// TwinCAT 3 PLC project Untitled2
// ProgramVersion: 3.1.4026.28
// libraries:
//   Tc2_Standard, * (Beckhoff Automation GmbH)
//   Tc2_System, * (Beckhoff Automation GmbH)
// project tree:
//   DUTs/ E_PackMLStates.TcDUT
//   / PlcTask.TcTTO
//   POUs/00_System/ MAIN.TcPOU
//   POUs/01_Unit/ FB_Unit.TcPOU
//   POUs/02_Equipment/01_Palletinvoer/ FB_Palletinvoer.TcPOU, ITF_Palletinvoer.TcIO
//   POUs/02_Equipment/02_Buffer2-4/ FB_Buffer2_4.TcPOU, ITF_Buffer2_4.TcIO
//   POUs/02_Equipment/03_Buffer5/ FB_Buffer5.TcPOU, ITF_Buffer5.TcIO
//   POUs/02_Equipment/04_Depalletizer/ FB_Depalletizer.TcPOU, ITF_Depalletizer.TcIO
//   POUs/02_Equipment/05_Banddepalletizer/ FB_Banddepalletizer.TcPOU, ITF_Banddepalletizer.TcIO
//   POUs/02_Equipment/06_Palletizer/ FB_Palletizer.TcPOU, ITF_Palletizer.TcIO
//   POUs/02_Equipment/07_Blikjesband/ FB_Blikjesband.TcPOU, ITF_Blikjesband.TcIO
//   POUs/02_Equipment/08_Besturing/ FB_Besturing.TcPOU, ITF_Besturing.TcIO
//   POUs/02_Equipment/ FB_Equipment.TcPOU
//   POUs/03_Control/ FB_Control.TcPOU
//   POUs/04_Management/Alarmmanager/ FB_Alarmmanager.TcPOU
//   POUs/04_Management/HMI/ FB_HMI.TcPOU
//   POUs/04_Management/Safety/ FB_Safety.TcPOU

CONFIGURATION Untitled2
    RESOURCE PLC ON TwinCAT3
        TASK PlcTask(INTERVAL := T#10ms, PRIORITY := 20);
        PROGRAM MAIN WITH PlcTask : MAIN;
    END_RESOURCE
END_CONFIGURATION

// ---- DUTs/E_PackMLStates.TcDUT
{attribute 'qualified_only'}
{attribute 'strict'}
{attribute 'to_string'}
TYPE E_PackMLStates :
(
	Idle := 0,
	Starting, 
	Execute, 
	Suspending, 
	Suspended, 
	Unsuspending, 
	Holding,
	Held,
	Unholding,
	Resetting,
	Aborting,
	Aborted, 
	Clearing,
	Stopping,
	Stopped
);
END_TYPE

// ---- POUs/02_Equipment/01_Palletinvoer/ITF_Palletinvoer.TcIO
INTERFACE ITF_Palletinvoer

METHOD Aborted : BOOL
VAR_INPUT
END_VAR
END_METHOD

METHOD Aborting : BOOL
VAR_INPUT
END_VAR
END_METHOD

METHOD Clearing : BOOL
VAR_INPUT
END_VAR
END_METHOD

METHOD Execute : BOOL
VAR_INPUT
END_VAR
END_METHOD

METHOD Held : BOOL
VAR_INPUT
END_VAR
END_METHOD

METHOD Holding : BOOL
VAR_INPUT
END_VAR
END_METHOD

METHOD Idle : BOOL
VAR_INPUT
END_VAR
END_METHOD

METHOD Resetting : BOOL
VAR_INPUT
END_VAR
END_METHOD

METHOD Starting : BOOL
VAR_INPUT
END_VAR
END_METHOD

METHOD Stopped : BOOL
VAR_INPUT
END_VAR
END_METHOD

METHOD Stopping : BOOL
VAR_INPUT
END_VAR
END_METHOD

METHOD Suspended : BOOL
VAR_INPUT
END_VAR
END_METHOD

METHOD Suspending : BOOL
VAR_INPUT
END_VAR
END_METHOD

METHOD Unholding : BOOL
VAR_INPUT
END_VAR
END_METHOD

METHOD Unsuspending : BOOL
VAR_INPUT
END_VAR
END_METHOD

END_INTERFACE

// ---- POUs/02_Equipment/02_Buffer2-4/ITF_Buffer2_4.TcIO
INTERFACE ITF_Buffer2_4

METHOD Aborted : BOOL
VAR_INPUT
END_VAR
END_METHOD

METHOD Aborting : BOOL
VAR_INPUT
END_VAR
END_METHOD

METHOD Clearing : BOOL
VAR_INPUT
END_VAR
END_METHOD

METHOD Execute : BOOL
VAR_INPUT
END_VAR
END_METHOD

METHOD Held : BOOL
VAR_INPUT
END_VAR
END_METHOD

METHOD Holding : BOOL
VAR_INPUT
END_VAR
END_METHOD

METHOD Idle : BOOL
VAR_INPUT
END_VAR
END_METHOD

METHOD Resetting : BOOL
VAR_INPUT
END_VAR
END_METHOD

METHOD Starting : BOOL
VAR_INPUT
END_VAR
END_METHOD

METHOD Stopped : BOOL
VAR_INPUT
END_VAR
END_METHOD

METHOD Stopping : BOOL
VAR_INPUT
END_VAR
END_METHOD

METHOD Suspended : BOOL
VAR_INPUT
END_VAR
END_METHOD

METHOD Suspending : BOOL
VAR_INPUT
END_VAR
END_METHOD

METHOD Unholding : BOOL
VAR_INPUT
END_VAR
END_METHOD

METHOD Unsuspending : BOOL
VAR_INPUT
END_VAR
END_METHOD

END_INTERFACE

// ---- POUs/02_Equipment/03_Buffer5/ITF_Buffer5.TcIO
INTERFACE ITF_Buffer5

METHOD Aborted : BOOL
VAR_INPUT
END_VAR
END_METHOD

METHOD Aborting : BOOL
VAR_INPUT
END_VAR
END_METHOD

METHOD Clearing : BOOL
VAR_INPUT
END_VAR
END_METHOD

METHOD Execute : BOOL
VAR_INPUT
END_VAR
END_METHOD

METHOD Held : BOOL
VAR_INPUT
END_VAR
END_METHOD

METHOD Holding : BOOL
VAR_INPUT
END_VAR
END_METHOD

METHOD Idle : BOOL
VAR_INPUT
END_VAR
END_METHOD

METHOD Resetting : BOOL
VAR_INPUT
END_VAR
END_METHOD

METHOD Starting : BOOL
VAR_INPUT
END_VAR
END_METHOD

METHOD Stopped : BOOL
VAR_INPUT
END_VAR
END_METHOD

METHOD Stopping : BOOL
VAR_INPUT
END_VAR
END_METHOD

METHOD Suspended : BOOL
VAR_INPUT
END_VAR
END_METHOD

METHOD Suspending : BOOL
VAR_INPUT
END_VAR
END_METHOD

METHOD Unholding : BOOL
VAR_INPUT
END_VAR
END_METHOD

METHOD Unsuspending : BOOL
VAR_INPUT
END_VAR
END_METHOD

END_INTERFACE

// ---- POUs/02_Equipment/04_Depalletizer/ITF_Depalletizer.TcIO
INTERFACE ITF_Depalletizer

METHOD Aborted : BOOL
VAR_INPUT
END_VAR
END_METHOD

METHOD Aborting : BOOL
VAR_INPUT
END_VAR
END_METHOD

METHOD Clearing : BOOL
VAR_INPUT
END_VAR
END_METHOD

METHOD Execute : BOOL
VAR_INPUT
END_VAR
END_METHOD

METHOD Held : BOOL
VAR_INPUT
END_VAR
END_METHOD

METHOD Holding : BOOL
VAR_INPUT
END_VAR
END_METHOD

METHOD Idle : BOOL
VAR_INPUT
END_VAR
END_METHOD

METHOD Resetting : BOOL
VAR_INPUT
END_VAR
END_METHOD

METHOD Starting : BOOL
VAR_INPUT
END_VAR
END_METHOD

METHOD Stopped : BOOL
VAR_INPUT
END_VAR
END_METHOD

METHOD Stopping : BOOL
VAR_INPUT
END_VAR
END_METHOD

METHOD Suspended : BOOL
VAR_INPUT
END_VAR
END_METHOD

METHOD Suspending : BOOL
VAR_INPUT
END_VAR
END_METHOD

METHOD Unholding : BOOL
VAR_INPUT
END_VAR
END_METHOD

METHOD Unsuspending : BOOL
VAR_INPUT
END_VAR
END_METHOD

END_INTERFACE

// ---- POUs/02_Equipment/05_Banddepalletizer/ITF_Banddepalletizer.TcIO
INTERFACE ITF_Banddepalletizer

METHOD Aborted : BOOL
VAR_INPUT
END_VAR
END_METHOD

METHOD Aborting : BOOL
VAR_INPUT
END_VAR
END_METHOD

METHOD Clearing : BOOL
VAR_INPUT
END_VAR
END_METHOD

METHOD Execute : BOOL
VAR_INPUT
END_VAR
END_METHOD

METHOD Held : BOOL
VAR_INPUT
END_VAR
END_METHOD

METHOD Holding : BOOL
VAR_INPUT
END_VAR
END_METHOD

METHOD Idle : BOOL
VAR_INPUT
END_VAR
END_METHOD

METHOD Resetting : BOOL
VAR_INPUT
END_VAR
END_METHOD

METHOD Starting : BOOL
VAR_INPUT
END_VAR
END_METHOD

METHOD Stopped : BOOL
VAR_INPUT
END_VAR
END_METHOD

METHOD Stopping : BOOL
VAR_INPUT
END_VAR
END_METHOD

METHOD Suspended : BOOL
VAR_INPUT
END_VAR
END_METHOD

METHOD Suspending : BOOL
VAR_INPUT
END_VAR
END_METHOD

METHOD Unholding : BOOL
VAR_INPUT
END_VAR
END_METHOD

METHOD Unsuspending : BOOL
VAR_INPUT
END_VAR
END_METHOD

END_INTERFACE

// ---- POUs/02_Equipment/06_Palletizer/ITF_Palletizer.TcIO
INTERFACE ITF_Palletizer

METHOD Aborted : BOOL
VAR_INPUT
END_VAR
END_METHOD

METHOD Aborting : BOOL
VAR_INPUT
END_VAR
END_METHOD

METHOD Clearing : BOOL
VAR_INPUT
END_VAR
END_METHOD

METHOD Execute : BOOL
VAR_INPUT
END_VAR
END_METHOD

METHOD Held : BOOL
VAR_INPUT
END_VAR
END_METHOD

METHOD Holding : BOOL
VAR_INPUT
END_VAR
END_METHOD

METHOD Idle : BOOL
VAR_INPUT
END_VAR
END_METHOD

METHOD Resetting : BOOL
VAR_INPUT
END_VAR
END_METHOD

METHOD Starting : BOOL
VAR_INPUT
END_VAR
END_METHOD

METHOD Stopped : BOOL
VAR_INPUT
END_VAR
END_METHOD

METHOD Stopping : BOOL
VAR_INPUT
END_VAR
END_METHOD

METHOD Suspended : BOOL
VAR_INPUT
END_VAR
END_METHOD

METHOD Suspending : BOOL
VAR_INPUT
END_VAR
END_METHOD

METHOD Unholding : BOOL
VAR_INPUT
END_VAR
END_METHOD

METHOD Unsuspending : BOOL
VAR_INPUT
END_VAR
END_METHOD

END_INTERFACE

// ---- POUs/02_Equipment/07_Blikjesband/ITF_Blikjesband.TcIO
INTERFACE ITF_Blikjesband

METHOD Aborted : BOOL
VAR_INPUT
END_VAR
END_METHOD

METHOD Aborting : BOOL
VAR_INPUT
END_VAR
END_METHOD

METHOD Clearing : BOOL
VAR_INPUT
END_VAR
END_METHOD

METHOD Execute : BOOL
VAR_INPUT
END_VAR
END_METHOD

METHOD Held : BOOL
VAR_INPUT
END_VAR
END_METHOD

METHOD Holding : BOOL
VAR_INPUT
END_VAR
END_METHOD

METHOD Idle : BOOL
VAR_INPUT
END_VAR
END_METHOD

METHOD Resetting : BOOL
VAR_INPUT
END_VAR
END_METHOD

METHOD Starting : BOOL
VAR_INPUT
END_VAR
END_METHOD

METHOD Stopped : BOOL
VAR_INPUT
END_VAR
END_METHOD

METHOD Stopping : BOOL
VAR_INPUT
END_VAR
END_METHOD

METHOD Suspended : BOOL
VAR_INPUT
END_VAR
END_METHOD

METHOD Suspending : BOOL
VAR_INPUT
END_VAR
END_METHOD

METHOD Unholding : BOOL
VAR_INPUT
END_VAR
END_METHOD

METHOD Unsuspending : BOOL
VAR_INPUT
END_VAR
END_METHOD

END_INTERFACE

// ---- POUs/02_Equipment/08_Besturing/ITF_Besturing.TcIO
INTERFACE ITF_Besturing

METHOD StatusLampGeel : BOOL
VAR_INPUT
END_VAR
END_METHOD

METHOD StatusLampGroen : BOOL
VAR_INPUT
END_VAR
END_METHOD

METHOD StatusLampRood : BOOL
VAR_INPUT
END_VAR
END_METHOD

END_INTERFACE

// ---- POUs/00_System/MAIN.TcPOU
PROGRAM MAIN
VAR
	test : BOOL;
END_VAR

// Klopt dit?

END_PROGRAM

// ---- POUs/01_Unit/FB_Unit.TcPOU
FUNCTION_BLOCK FB_Unit
VAR_INPUT
END_VAR
VAR_OUTPUT
END_VAR
VAR
END_VAR

END_FUNCTION_BLOCK

// ---- POUs/02_Equipment/01_Palletinvoer/FB_Palletinvoer.TcPOU
FUNCTION_BLOCK FB_Palletinvoer IMPLEMENTS ITF_Palletinvoer
VAR_INPUT
END_VAR
VAR_OUTPUT
END_VAR
VAR
END_VAR

{warning 'Add method implementation '}
METHOD Aborted : BOOL
END_METHOD

{warning 'Add method implementation '}
METHOD Aborting : BOOL
END_METHOD

{warning 'Add method implementation '}
METHOD Clearing : BOOL
END_METHOD

{warning 'Add method implementation '}
METHOD Execute : BOOL
END_METHOD

{warning 'Add method implementation '}
METHOD Held : BOOL
END_METHOD

{warning 'Add method implementation '}
METHOD Holding : BOOL
END_METHOD

{warning 'Add method implementation '}
METHOD Idle : BOOL
END_METHOD

{warning 'Add method implementation '}
METHOD Resetting : BOOL
END_METHOD

{warning 'Add method implementation '}
METHOD Starting : BOOL
END_METHOD

{warning 'Add method implementation '}
METHOD Stopped : BOOL
END_METHOD

{warning 'Add method implementation '}
METHOD Stopping : BOOL
END_METHOD

{warning 'Add method implementation '}
METHOD Suspended : BOOL
END_METHOD

{warning 'Add method implementation '}
METHOD Suspending : BOOL
END_METHOD

{warning 'Add method implementation '}
METHOD Unholding : BOOL
END_METHOD

{warning 'Add method implementation '}
METHOD Unsuspending : BOOL
END_METHOD

END_FUNCTION_BLOCK

// ---- POUs/02_Equipment/02_Buffer2-4/FB_Buffer2_4.TcPOU
FUNCTION_BLOCK FB_Buffer2_4 IMPLEMENTS ITF_Buffer2_4
VAR_INPUT
END_VAR
VAR_OUTPUT
END_VAR
VAR
END_VAR

{warning 'Add method implementation '}
METHOD Aborted : BOOL
END_METHOD

{warning 'Add method implementation '}
METHOD Aborting : BOOL
END_METHOD

{warning 'Add method implementation '}
METHOD Clearing : BOOL
END_METHOD

{warning 'Add method implementation '}
METHOD Execute : BOOL
END_METHOD

{warning 'Add method implementation '}
METHOD Held : BOOL
END_METHOD

{warning 'Add method implementation '}
METHOD Holding : BOOL
END_METHOD

{warning 'Add method implementation '}
METHOD Idle : BOOL
END_METHOD

{warning 'Add method implementation '}
METHOD Resetting : BOOL
END_METHOD

{warning 'Add method implementation '}
METHOD Starting : BOOL
END_METHOD

{warning 'Add method implementation '}
METHOD Stopped : BOOL
END_METHOD

{warning 'Add method implementation '}
METHOD Stopping : BOOL
END_METHOD

{warning 'Add method implementation '}
METHOD Suspended : BOOL
END_METHOD

{warning 'Add method implementation '}
METHOD Suspending : BOOL
END_METHOD

{warning 'Add method implementation '}
METHOD Unholding : BOOL
END_METHOD

{warning 'Add method implementation '}
METHOD Unsuspending : BOOL
END_METHOD

END_FUNCTION_BLOCK

// ---- POUs/02_Equipment/03_Buffer5/FB_Buffer5.TcPOU
FUNCTION_BLOCK FB_Buffer5 IMPLEMENTS ITF_Buffer5
VAR_INPUT
END_VAR
VAR_OUTPUT
END_VAR
VAR
END_VAR

{warning 'Add method implementation '}
METHOD Aborted : BOOL
END_METHOD

{warning 'Add method implementation '}
METHOD Aborting : BOOL
END_METHOD

{warning 'Add method implementation '}
METHOD Clearing : BOOL
END_METHOD

{warning 'Add method implementation '}
METHOD Execute : BOOL
END_METHOD

{warning 'Add method implementation '}
METHOD Held : BOOL
END_METHOD

{warning 'Add method implementation '}
METHOD Holding : BOOL
END_METHOD

{warning 'Add method implementation '}
METHOD Idle : BOOL
END_METHOD

{warning 'Add method implementation '}
METHOD Resetting : BOOL
END_METHOD

{warning 'Add method implementation '}
METHOD Starting : BOOL
END_METHOD

{warning 'Add method implementation '}
METHOD Stopped : BOOL
END_METHOD

{warning 'Add method implementation '}
METHOD Stopping : BOOL
END_METHOD

{warning 'Add method implementation '}
METHOD Suspended : BOOL
END_METHOD

{warning 'Add method implementation '}
METHOD Suspending : BOOL
END_METHOD

{warning 'Add method implementation '}
METHOD Unholding : BOOL
END_METHOD

{warning 'Add method implementation '}
METHOD Unsuspending : BOOL
END_METHOD

END_FUNCTION_BLOCK

// ---- POUs/02_Equipment/04_Depalletizer/FB_Depalletizer.TcPOU
FUNCTION_BLOCK FB_Depalletizer IMPLEMENTS ITF_Depalletizer
VAR_INPUT
END_VAR
VAR_OUTPUT
END_VAR
VAR
END_VAR

{warning 'Add method implementation '}
METHOD Aborted : BOOL
END_METHOD

{warning 'Add method implementation '}
METHOD Aborting : BOOL
END_METHOD

{warning 'Add method implementation '}
METHOD Clearing : BOOL
END_METHOD

{warning 'Add method implementation '}
METHOD Execute : BOOL
END_METHOD

{warning 'Add method implementation '}
METHOD Held : BOOL
END_METHOD

{warning 'Add method implementation '}
METHOD Holding : BOOL
END_METHOD

{warning 'Add method implementation '}
METHOD Idle : BOOL
END_METHOD

{warning 'Add method implementation '}
METHOD Resetting : BOOL
END_METHOD

{warning 'Add method implementation '}
METHOD Starting : BOOL
END_METHOD

{warning 'Add method implementation '}
METHOD Stopped : BOOL
END_METHOD

{warning 'Add method implementation '}
METHOD Stopping : BOOL
END_METHOD

{warning 'Add method implementation '}
METHOD Suspended : BOOL
END_METHOD

{warning 'Add method implementation '}
METHOD Suspending : BOOL
END_METHOD

{warning 'Add method implementation '}
METHOD Unholding : BOOL
END_METHOD

{warning 'Add method implementation '}
METHOD Unsuspending : BOOL
END_METHOD

END_FUNCTION_BLOCK

// ---- POUs/02_Equipment/05_Banddepalletizer/FB_Banddepalletizer.TcPOU
FUNCTION_BLOCK FB_Banddepalletizer IMPLEMENTS ITF_Banddepalletizer
VAR_INPUT
END_VAR
VAR_OUTPUT
END_VAR
VAR
END_VAR

{warning 'Add method implementation '}
METHOD Aborted : BOOL
END_METHOD

{warning 'Add method implementation '}
METHOD Aborting : BOOL
END_METHOD

{warning 'Add method implementation '}
METHOD Clearing : BOOL
END_METHOD

{warning 'Add method implementation '}
METHOD Execute : BOOL
END_METHOD

{warning 'Add method implementation '}
METHOD Held : BOOL
END_METHOD

{warning 'Add method implementation '}
METHOD Holding : BOOL
END_METHOD

{warning 'Add method implementation '}
METHOD Idle : BOOL
END_METHOD

{warning 'Add method implementation '}
METHOD Resetting : BOOL
END_METHOD

{warning 'Add method implementation '}
METHOD Starting : BOOL
END_METHOD

{warning 'Add method implementation '}
METHOD Stopped : BOOL
END_METHOD

{warning 'Add method implementation '}
METHOD Stopping : BOOL
END_METHOD

{warning 'Add method implementation '}
METHOD Suspended : BOOL
END_METHOD

{warning 'Add method implementation '}
METHOD Suspending : BOOL
END_METHOD

{warning 'Add method implementation '}
METHOD Unholding : BOOL
END_METHOD

{warning 'Add method implementation '}
METHOD Unsuspending : BOOL
END_METHOD

END_FUNCTION_BLOCK

// ---- POUs/02_Equipment/06_Palletizer/FB_Palletizer.TcPOU
FUNCTION_BLOCK FB_Palletizer IMPLEMENTS ITF_Palletizer
VAR_INPUT
END_VAR
VAR_OUTPUT
END_VAR
VAR
END_VAR

{warning 'Add method implementation '}
METHOD Aborted : BOOL
END_METHOD

{warning 'Add method implementation '}
METHOD Aborting : BOOL
END_METHOD

{warning 'Add method implementation '}
METHOD Clearing : BOOL
END_METHOD

{warning 'Add method implementation '}
METHOD Execute : BOOL
END_METHOD

{warning 'Add method implementation '}
METHOD Held : BOOL
END_METHOD

{warning 'Add method implementation '}
METHOD Holding : BOOL
END_METHOD

{warning 'Add method implementation '}
METHOD Idle : BOOL
END_METHOD

{warning 'Add method implementation '}
METHOD Resetting : BOOL
END_METHOD

{warning 'Add method implementation '}
METHOD Starting : BOOL
END_METHOD

{warning 'Add method implementation '}
METHOD Stopped : BOOL
END_METHOD

{warning 'Add method implementation '}
METHOD Stopping : BOOL
END_METHOD

{warning 'Add method implementation '}
METHOD Suspended : BOOL
END_METHOD

{warning 'Add method implementation '}
METHOD Suspending : BOOL
END_METHOD

{warning 'Add method implementation '}
METHOD Unholding : BOOL
END_METHOD

{warning 'Add method implementation '}
METHOD Unsuspending : BOOL
END_METHOD

END_FUNCTION_BLOCK

// ---- POUs/02_Equipment/07_Blikjesband/FB_Blikjesband.TcPOU
FUNCTION_BLOCK FB_Blikjesband IMPLEMENTS ITF_Blikjesband
VAR_INPUT
END_VAR
VAR_OUTPUT
END_VAR
VAR
END_VAR

{warning 'Add method implementation '}
METHOD Aborted : BOOL
END_METHOD

{warning 'Add method implementation '}
METHOD Aborting : BOOL
END_METHOD

{warning 'Add method implementation '}
METHOD Clearing : BOOL
END_METHOD

{warning 'Add method implementation '}
METHOD Execute : BOOL
END_METHOD

{warning 'Add method implementation '}
METHOD Held : BOOL
END_METHOD

{warning 'Add method implementation '}
METHOD Holding : BOOL
END_METHOD

{warning 'Add method implementation '}
METHOD Idle : BOOL
END_METHOD

{warning 'Add method implementation '}
METHOD Resetting : BOOL
END_METHOD

{warning 'Add method implementation '}
METHOD Starting : BOOL
END_METHOD

{warning 'Add method implementation '}
METHOD Stopped : BOOL
END_METHOD

{warning 'Add method implementation '}
METHOD Stopping : BOOL
END_METHOD

{warning 'Add method implementation '}
METHOD Suspended : BOOL
END_METHOD

{warning 'Add method implementation '}
METHOD Suspending : BOOL
END_METHOD

{warning 'Add method implementation '}
METHOD Unholding : BOOL
END_METHOD

{warning 'Add method implementation '}
METHOD Unsuspending : BOOL
END_METHOD

END_FUNCTION_BLOCK

// ---- POUs/02_Equipment/08_Besturing/FB_Besturing.TcPOU
FUNCTION_BLOCK FB_Besturing IMPLEMENTS ITF_Besturing
VAR_INPUT
END_VAR
VAR_OUTPUT
END_VAR
VAR
END_VAR

{warning 'Add method implementation '}
METHOD StatusLampGeel : BOOL
END_METHOD

{warning 'Add method implementation '}
METHOD StatusLampGroen : BOOL
END_METHOD

{warning 'Add method implementation '}
METHOD StatusLampRood : BOOL
END_METHOD

END_FUNCTION_BLOCK

// ---- POUs/02_Equipment/FB_Equipment.TcPOU
FUNCTION_BLOCK FB_Equipment
VAR_INPUT
END_VAR
VAR_OUTPUT
END_VAR
VAR
END_VAR

END_FUNCTION_BLOCK

// ---- POUs/03_Control/FB_Control.TcPOU
FUNCTION_BLOCK FB_Control
VAR_INPUT
END_VAR
VAR_OUTPUT
END_VAR
VAR
END_VAR

END_FUNCTION_BLOCK

// ---- POUs/04_Management/Alarmmanager/FB_Alarmmanager.TcPOU
FUNCTION_BLOCK FB_Alarmmanager
VAR_INPUT
END_VAR
VAR_OUTPUT
END_VAR
VAR
END_VAR

END_FUNCTION_BLOCK

// ---- POUs/04_Management/HMI/FB_HMI.TcPOU
FUNCTION_BLOCK FB_HMI
VAR_INPUT
END_VAR
VAR_OUTPUT
END_VAR
VAR
END_VAR

END_FUNCTION_BLOCK

// ---- POUs/04_Management/Safety/FB_Safety.TcPOU
FUNCTION_BLOCK FB_Safety
VAR_INPUT
END_VAR
VAR_OUTPUT
END_VAR
VAR
END_VAR

END_FUNCTION_BLOCK
